Fanuc KAREL source: KA00108.KL

PROGRAM KA00108
%NOLOCKGROUP
VAR
  SRC: VECTOR
  DST: ARRAY[2] OF SHORT
BEGIN
  SRC.X = 1.0
  DST[1] = SRC
END KA00108
